Staubli VAL3: main.pgx

program main()
begin
  close(tCurrentTool)
  pPointRx.config.shoulder = lefty
  pPointRx.config.elbow = epositive
  pPointRx.config.wrist = wpositive
  pPointRx2.config.shoulder = lefty
  pPointRx2.config.elbow = epositive
  pPointRx2.config.wrist = wpositive
  mCurrentSpeed.tvel = 100.00
  mCurrentSpeed.blend = joint
  mCurrentSpeed.reach = 0.010
  mCurrentSpeed.leave = 0.010
  // Program JointTargets start
  // Program generated by VerticalBot Studio for Staubli RX160 on 25/10/2026 12:00:00
  // Using nominal kinematics.
  call MoveJoint(10.00000,20.00000,90.00000,30.00000,45.00000,60.00000)
  // Linear movement using joint targets is not supported. Change the target type to cartesian or use a joint movement.
  call MoveJoint(18.00000,24.00000,90.00000,30.00000,45.00000,60.00000)
  call MoveLine(1023.000,-205.063,905.909,-149.902,32.793,-96.693)
  // Linear movement using joint targets is not supported. Change the target type to cartesian or use a joint movement.
  mCurrentSpeed.reach = 5.000
  mCurrentSpeed.leave = 5.000
  call MoveJoint(10.00000,20.00000,90.00000,30.00000,45.00000,60.00000)
  // Linear movement using joint targets is not supported. Change the target type to cartesian or use a joint movement.
  call MoveJoint(18.00000,24.00000,90.00000,30.00000,45.00000,60.00000)
  call MoveLine(1023.000,-205.063,905.909,-149.902,32.793,-96.693)
  // Linear movement using joint targets is not supported. Change the target type to cartesian or use a joint movement.
  mCurrentSpeed.reach = -1.000
  mCurrentSpeed.leave = -1.000
  call MoveJoint(10.00000,20.00000,90.00000,30.00000,45.00000,60.00000)

  waitEndMove()
  // Program JointTargets end

end
